Fanuc KAREL source: kc00061.KL

-- PROVISIONAL review KL for V940-1; original PC SHA256 51b8773c171b182eeeaca20ff90436fbb9f948112236ef611efba7a5623bf1df
-- Incomplete behavior may be omitted. Consult companion uncertainty JSON. Do not deploy.
PROGRAM KC00061
%NOLOCKGROUP
BEGIN
  -- V9_ZERO_TABLE_METADATA_HINT layout=0002_ascii; no indexed target words; source/name/runtime held
  -- UNRESOLVED_PC offsets 5-37; opcodes 27,27,9D,27,9D,22,1C,22,AA,23
  -- UNRESOLVED_PC offsets 42-46; opcodes 7F
END KC00061
